(* CODESYS project SysParBuggy.xml

Project tree, tasks and I/O mapping:
  visualisation SysParBuggy
*)

// /SysParBuggy
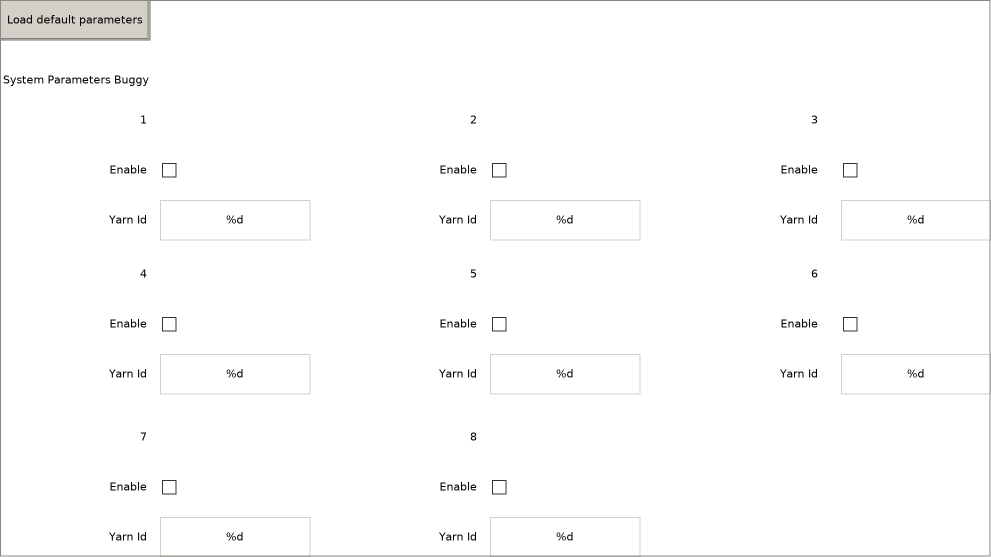
VISUALIZATION SysParBuggy  // 991x557
    Button (0,0 150x40), "Load default parameters"
        tap PRG_VisuTask_10ms._fbParametersCtrl._btnLoadDefaultParameters.xbtn
    Label (0,60 300x40), "System Parameters Buggy"
    Label (0,200 150x40), "Yarn Id"
    Textfield (160,200 150x40), "%d", text variable: PersistentVars.scYarnStorages.ascYarnStorage[1].iYarnType
        OnMouseUp: write the text variable via Default
    Label (0,150 150x40), "Enable"
    Checkbox (160,150 40x40), variable: PersistentVars.scYarnStorages.ascYarnStorage[1].xEnabled
    Label (0,100 150x40), "1"
    Label (671,200 150x40), "Yarn Id"
    Textfield (841,200 150x40), "%d", text variable: PersistentVars.scYarnStorages.ascYarnStorage[3].iYarnType
        OnMouseUp: write the text variable via Default
    Label (671,150 150x40), "Enable"
    Checkbox (841,150 40x40), variable: PersistentVars.scYarnStorages.ascYarnStorage[3].xEnabled
    Label (671,100 150x40), "3"
    Label (330,200 150x40), "Yarn Id"
    Textfield (490,200 150x40), "%d", text variable: PersistentVars.scYarnStorages.ascYarnStorage[2].iYarnType
        OnMouseUp: write the text variable via Default
    Label (330,150 150x40), "Enable"
    Checkbox (490,150 40x40), variable: PersistentVars.scYarnStorages.ascYarnStorage[2].xEnabled
    Label (330,100 150x40), "2"
    Label (0,354 150x40), "Yarn Id"
    Textfield (160,354 150x40), "%d", text variable: PersistentVars.scYarnStorages.ascYarnStorage[4].iYarnType
        OnMouseUp: write the text variable via Default
    Label (0,304 150x40), "Enable"
    Checkbox (160,304 40x40), variable: PersistentVars.scYarnStorages.ascYarnStorage[4].xEnabled
    Label (0,254 150x40), "4"
    Label (330,354 150x40), "Yarn Id"
    Textfield (490,354 150x40), "%d", text variable: PersistentVars.scYarnStorages.ascYarnStorage[5].iYarnType
        OnMouseUp: write the text variable via Default
    Label (330,304 150x40), "Enable"
    Checkbox (490,304 40x40), variable: PersistentVars.scYarnStorages.ascYarnStorage[5].xEnabled
    Label (330,254 150x40), "5"
    Label (671,354 150x40), "Yarn Id"
    Textfield (841,354 150x40), "%d", text variable: PersistentVars.scYarnStorages.ascYarnStorage[6].iYarnType
        OnMouseUp: write the text variable via Default
    Label (671,304 150x40), "Enable"
    Checkbox (841,304 40x40), variable: PersistentVars.scYarnStorages.ascYarnStorage[6].xEnabled
    Label (671,254 150x40), "6"
    Label (0,517 150x40), "Yarn Id"
    Textfield (160,517 150x40), "%d", text variable: PersistentVars.scYarnStorages.ascYarnStorage[7].iYarnType
        OnMouseUp: write the text variable via Default
    Label (0,467 150x40), "Enable"
    Checkbox (160,467 40x40), variable: PersistentVars.scYarnStorages.ascYarnStorage[7].xEnabled
    Label (0,417 150x40), "7"
    Label (330,517 150x40), "Yarn Id"
    Textfield (490,517 150x40), "%d", text variable: PersistentVars.scYarnStorages.ascYarnStorage[8].iYarnType
        OnMouseUp: write the text variable via Default
    Label (330,467 150x40), "Enable"
    Checkbox (490,467 40x40), variable: PersistentVars.scYarnStorages.ascYarnStorage[8].xEnabled
    Label (330,417 150x40), "8"
END_VISUALIZATION
